(* IEC 61131-3 sources: SafePLC-Gen-Evaluation/Evaluation Results/butane/run_04, 2 files *)

(* ---- io_declarations.st ---- *)
(* ==================================================  *)
(* PLC I/O Variable Declarations — CODESYS 3.5  *)
(* Generated by SafePLC-Gen Multimodal  *)
(* ==================================================  *)

VAR_GLOBAL
    (* --- Analog Inputs ---  *)
    TI_2909_Raw                  AT %IW0       : INT := 0;    (* TI-2909 — Temperature indicator on process inlet l  *)
    TI_2917_Raw                  AT %IW2       : INT := 0;    (* TI-2917 — Temperature indicator high-high (HH), fa  *)
    TT_2909_Raw                  AT %IW4       : INT := 0;    (* TT-2909 — Temperature transmitter on process line,  *)
    TT_2911_Raw                  AT %IW6       : INT := 0;    (* TT-2911 — Temperature transmitter on process outle  *)
    TT_2917_Raw                  AT %IW8       : INT := 0;    (* TT-2917 — Temperature transmitter on heating mediu  *)
    XI_2901A_Raw                 AT %IW10      : INT := 0;    (* XI-2901A — Status indicator AVAILABLE for motor/fan  *)
    XI_2901B_Raw                 AT %IW12      : INT := 0;    (* XI-2901B — Status indicator AVAILABLE for motor/fan  *)
    (* --- Analog Outputs ---  *)
    KV_2904_Out                  AT %QW0       : INT := 0;    (* KV-2904 — Actuated valve on inlet process line, fa  *)
    (* --- Digital Inputs ---  *)
    ESD_3200                     AT %IX0.0     : BOOL := FALSE;    (* ESD-3200 — Emergency shutdown device/input, appears  *)
    HS_2901A                     AT %IX0.1     : BOOL := FALSE;    (* HS-2901A — Hand switch for motor/fan A control. Pan  *)
    HS_2901A1                    AT %IX0.2     : BOOL := FALSE;    (* HS-2901A1 — Hand switch LOCAL/REMOTE selector for mo  *)
    HS_2901A2                    AT %IX0.3     : BOOL := FALSE;    (* HS-2901A2 — Hand switch STOP/START for motor A at MC  *)
    HS_2901B                     AT %IX0.4     : BOOL := FALSE;    (* HS-2901B — Hand switch for motor/fan B control. Pan  *)
    HS_2901B1                    AT %IX0.5     : BOOL := FALSE;    (* HS-2901B1 — Hand switch LOCAL/REMOTE selector for mo  *)
    HS_2901B2                    AT %IX0.6     : BOOL := FALSE;    (* HS-2901B2 — Hand switch STOP/START for motor B at MC  *)
    HS_EMERGENCY_STOP_A_2901A    AT %IX0.7     : BOOL := FALSE;    (* HS-EMERGENCY-STOP-A-2901A — Emergency stop hand switch for motor A,   *)
    HS_EMERGENCY_STOP_B_2901B    AT %IX1.0     : BOOL := FALSE;    (* HS-EMERGENCY-STOP-B-2901B — Emergency stop hand switch for motor B,   *)
    HS_START_STOP_A_2901A        AT %IX1.1     : BOOL := FALSE;    (* HS-START-STOP-A-2901A — Field/local hand switch START/STOP for m  *)
    HS_START_STOP_B_2901B        AT %IX1.2     : BOOL := FALSE;    (* HS-START-STOP-B-2901B — Field/local hand switch START/STOP for m  *)
    PSD_2917                     AT %IX1.3     : BOOL := FALSE;    (* PSD-2917 — Pressure/Temperature shutdown device (PS  *)
    VSHH_2901A                   AT %IX1.4     : BOOL := FALSE;    (* VSHH-2901A — Vibration switch high-high on fan/motor   *)
    VSHH_2901B                   AT %IX1.5     : BOOL := FALSE;    (* VSHH-2901B — Vibration switch high-high on fan/motor   *)
END_VAR

(* ---- generated_code.st ---- *)
(* Generated by SafePLC-Gen Multimodal — CODESYS 3.5 *)
(* IEC 61131-3 Structured Text *)
(* Date: 2026-04-25T12:15:34.199960 *)

PROGRAM PRG_Compressor_2901

VAR
    TI_2909_Raw                  AT %IW0       : INT := 0;
    TI_2917_Raw                  AT %IW2       : INT := 0;
    TT_2909_Raw                  AT %IW4       : INT := 0;
    TT_2911_Raw                  AT %IW6       : INT := 0;
    TT_2917_Raw                  AT %IW8       : INT := 0;
    XI_2901A_Raw                 AT %IW10      : INT := 0;
    XI_2901B_Raw                 AT %IW12      : INT := 0;
    KV_2904_Out                  AT %QW0       : INT := 0;
    ESD_3200                     AT %IX0.0     : BOOL := FALSE;
    HS_2901A                     AT %IX0.1     : BOOL := FALSE;
    HS_2901A1                    AT %IX0.2     : BOOL := FALSE;
    HS_2901A2                    AT %IX0.3     : BOOL := FALSE;
    HS_2901B                     AT %IX0.4     : BOOL := FALSE;
    HS_2901B1                    AT %IX0.5     : BOOL := FALSE;
    HS_2901B2                    AT %IX0.6     : BOOL := FALSE;
    HS_EMERGENCY_STOP_A_2901A    AT %IX0.7     : BOOL := FALSE;
    HS_EMERGENCY_STOP_B_2901B    AT %IX1.0     : BOOL := FALSE;
    HS_START_STOP_A_2901A        AT %IX1.1     : BOOL := FALSE;
    HS_START_STOP_B_2901B        AT %IX1.2     : BOOL := FALSE;
    PSD_2917                     AT %IX1.3     : BOOL := FALSE;
    VSHH_2901A                   AT %IX1.4     : BOOL := FALSE;
    VSHH_2901B                   AT %IX1.5     : BOOL := FALSE;
    ESTOP                        AT %IX2.0     : BOOL := FALSE;
    MANUAL_RESET                 AT %IX2.1     : BOOL := FALSE;
    MCC_A_Out                    AT %QX0.0     : BOOL := FALSE;
    MCC_B_Out                    AT %QX0.1     : BOOL := FALSE;
    PSD_2917_Out                 AT %QX0.2     : BOOL := FALSE;
    MCC_A_and_MCC_B_Out          AT %QX0.3     : BOOL := FALSE;
END_VAR

VAR
    TI_2909_Scaled               : REAL := 0.0;
    TT_2909_Scaled               : REAL := 0.0;
    TT_2911_Scaled               : REAL := 0.0;
    TT_2917_Scaled               : REAL := 0.0;
    TI_2917_Scaled               : REAL := 0.0;
    XI_2901A_Scaled              : REAL := 0.0;
    XI_2901B_Scaled              : REAL := 0.0;

    TI_2909_HH_SP                : REAL := 120.0;
    TI_2909_H_SP                 : REAL := 110.0;
    TI_2909_L_SP                 : REAL := 10.0;
    TI_2909_LL_SP                : REAL := 5.0;
    TI_2909_Deadband             : REAL := 2.0;
    TI_2909_HH                   : BOOL := FALSE;
    TI_2909_H                    : BOOL := FALSE;
    TI_2909_L                    : BOOL := FALSE;
    TI_2909_LL                   : BOOL := FALSE;
    TI_2909_HH_Latch             : SR := (S1 := FALSE, R := FALSE, Q1 := FALSE);
    TI_2909_LL_Latch             : SR := (S1 := FALSE, R := FALSE, Q1 := FALSE);
    TI_2909_HH_Ack               : BOOL := FALSE;
    TI_2909_LL_Ack               : BOOL := FALSE;

    TT_2909_HH_SP                : REAL := 120.0;
    TT_2909_H_SP                 : REAL := 110.0;
    TT_2909_L_SP                 : REAL := 10.0;
    TT_2909_LL_SP                : REAL := 5.0;
    TT_2909_Deadband             : REAL := 2.0;
    TT_2909_HH                   : BOOL := FALSE;
    TT_2909_H                    : BOOL := FALSE;
    TT_2909_L                    : BOOL := FALSE;
    TT_2909_LL                   : BOOL := FALSE;
    TT_2909_HH_Latch             : SR := (S1 := FALSE, R := FALSE, Q1 := FALSE);
    TT_2909_LL_Latch             : SR := (S1 := FALSE, R := FALSE, Q1 := FALSE);
    TT_2909_HH_Ack               : BOOL := FALSE;
    TT_2909_LL_Ack               : BOOL := FALSE;

    TT_2911_HH_SP                : REAL := 120.0;
    TT_2911_H_SP                 : REAL := 110.0;
    TT_2911_L_SP                 : REAL := 10.0;
    TT_2911_LL_SP                : REAL := 5.0;
    TT_2911_Deadband             : REAL := 2.0;
    TT_2911_HH                   : BOOL := FALSE;
    TT_2911_H                    : BOOL := FALSE;
    TT_2911_L                    : BOOL := FALSE;
    TT_2911_LL                   : BOOL := FALSE;
    TT_2911_HH_Latch             : SR := (S1 := FALSE, R := FALSE, Q1 := FALSE);
    TT_2911_LL_Latch             : SR := (S1 := FALSE, R := FALSE, Q1 := FALSE);
    TT_2911_HH_Ack               : BOOL := FALSE;
    TT_2911_LL_Ack               : BOOL := FALSE;

    TIC_2911_SP                  : REAL := 60.0;
    TIC_2911_Kp                  : REAL := 1.5;
    TIC_2911_Ki                  : REAL := 0.05;
    TIC_2911_Error               : REAL := 0.0;
    TIC_2911_Integral            : REAL := 0.0;
    TIC_2911_Output              : REAL := 0.0;

    TT_2917_HH_SP                : REAL := 130.0;
    TT_2917_H_SP                 : REAL := 120.0;
    TT_2917_L_SP                 : REAL := 10.0;
    TT_2917_LL_SP                : REAL := 5.0;
    TT_2917_Deadband             : REAL := 2.0;
    TT_2917_HH                   : BOOL := FALSE;
    TT_2917_H                    : BOOL := FALSE;
    TT_2917_L                    : BOOL := FALSE;
    TT_2917_LL                   : BOOL := FALSE;
    TT_2917_HH_Latch             : SR := (S1 := FALSE, R := FALSE, Q1 := FALSE);
    TT_2917_LL_Latch             : SR := (S1 := FALSE, R := FALSE, Q1 := FALSE);
    TT_2917_HH_Ack               : BOOL := FALSE;
    TT_2917_LL_Ack               : BOOL := FALSE;

    TI_2917_HH_SP                : REAL := 130.0;
    TI_2917_H_SP                 : REAL := 120.0;
    TI_2917_L_SP                 : REAL := 10.0;
    TI_2917_LL_SP                : REAL := 5.0;
    TI_2917_Deadband             : REAL := 2.0;
    TI_2917_HH                   : BOOL := FALSE;
    TI_2917_H                    : BOOL := FALSE;
    TI_2917_L                    : BOOL := FALSE;
    TI_2917_LL                   : BOOL := FALSE;
    TI_2917_HH_Latch             : SR := (S1 := FALSE, R := FALSE, Q1 := FALSE);
    TI_2917_LL_Latch             : SR := (S1 := FALSE, R := FALSE, Q1 := FALSE);
    TI_2917_HH_Ack               : BOOL := FALSE;
    TI_2917_LL_Ack               : BOOL := FALSE;

    XI_2901A_HH_SP               : REAL := 90.0;
    XI_2901A_H_SP                : REAL := 80.0;
    XI_2901A_L_SP                : REAL := 10.0;
    XI_2901A_LL_SP               : REAL := 5.0;
    XI_2901A_Deadband            : REAL := 2.0;
    XI_2901A_HH                  : BOOL := FALSE;
    XI_2901A_H                   : BOOL := FALSE;
    XI_2901A_L                   : BOOL := FALSE;
    XI_2901A_LL                  : BOOL := FALSE;
    XI_2901A_HH_Latch            : SR := (S1 := FALSE, R := FALSE, Q1 := FALSE);
    XI_2901A_LL_Latch            : SR := (S1 := FALSE, R := FALSE, Q1 := FALSE);
    XI_2901A_HH_Ack              : BOOL := FALSE;
    XI_2901A_LL_Ack              : BOOL := FALSE;

    XI_2901B_HH_SP               : REAL := 90.0;
    XI_2901B_H_SP                : REAL := 80.0;
    XI_2901B_L_SP                : REAL := 10.0;
    XI_2901B_LL_SP               : REAL := 5.0;
    XI_2901B_Deadband            : REAL := 2.0;
    XI_2901B_HH                  : BOOL := FALSE;
    XI_2901B_H                   : BOOL := FALSE;
    XI_2901B_L                   : BOOL := FALSE;
    XI_2901B_LL                  : BOOL := FALSE;
    XI_2901B_HH_Latch            : SR := (S1 := FALSE, R := FALSE, Q1 := FALSE);
    XI_2901B_LL_Latch            : SR := (S1 := FALSE, R := FALSE, Q1 := FALSE);
    XI_2901B_HH_Ack              : BOOL := FALSE;
    XI_2901B_LL_Ack              : BOOL := FALSE;

    LOOP_2917_TRIP               : BOOL := FALSE;
    LOOP_2901A_TRIP              : BOOL := FALSE;
    LOOP_2901B_TRIP              : BOOL := FALSE;
    LOOP_3200_TRIP               : BOOL := FALSE;

    TT_2917_HH_Trip              : BOOL := FALSE;
    TT_2917_LL_Trip              : BOOL := FALSE;
    VSHH_2901A_HH                : BOOL := FALSE;
    VSHH_2901A_LL                : BOOL := FALSE;
    VSHH_2901B_HH                : BOOL := FALSE;
    VSHH_2901B_LL                : BOOL := FALSE;
    ESD_3200_HH                  : BOOL := FALSE;
    ESD_3200_LL                  : BOOL := FALSE;

    SAFE_STATE                   : BOOL := FALSE;

    MotorA_LocalMode             : BOOL := FALSE;
    MotorA_StartCmd              : BOOL := FALSE;
    MotorA_StopCmd               : BOOL := FALSE;
    MotorA_Run                   : BOOL := FALSE;
    MotorA_Latch                 : SR := (S1 := FALSE, R := FALSE, Q1 := FALSE);

    MotorB_LocalMode             : BOOL := FALSE;
    MotorB_StartCmd              : BOOL := FALSE;
    MotorB_StopCmd               : BOOL := FALSE;
    MotorB_Run                   : BOOL := FALSE;
    MotorB_Latch                 : SR := (S1 := FALSE, R := FALSE, Q1 := FALSE);

    StartupDelay                 : TON := (IN := FALSE, PT := T#3S);

    System_Alarm                 : BOOL := FALSE;
    FirstScan                    : BOOL := TRUE;
END_VAR

IF FirstScan THEN
    LOOP_2917_TRIP       := TRUE;
    LOOP_2901A_TRIP      := TRUE;
    LOOP_2901B_TRIP      := TRUE;
    LOOP_3200_TRIP       := TRUE;
    SAFE_STATE           := TRUE;
    KV_2904_Out          := 6554;
    MCC_A_Out            := FALSE;
    MCC_B_Out            := FALSE;
    PSD_2917_Out         := FALSE;
    MCC_A_and_MCC_B_Out  := FALSE;
    TIC_2911_Integral    := 0.0;
    FirstScan            := FALSE;
    RETURN;
END_IF;

TI_2909_Scaled  := ((INT_TO_REAL(TI_2909_Raw)  - 6554.0) / (32767.0 - 6554.0)) * 150.0;
TT_2909_Scaled  := ((INT_TO_REAL(TT_2909_Raw)  - 6554.0) / (32767.0 - 6554.0)) * 150.0;
TT_2911_Scaled  := ((INT_TO_REAL(TT_2911_Raw)  - 6554.0) / (32767.0 - 6554.0)) * 150.0;
TT_2917_Scaled  := ((INT_TO_REAL(TT_2917_Raw)  - 6554.0) / (32767.0 - 6554.0)) * 150.0;
TI_2917_Scaled  := ((INT_TO_REAL(TI_2917_Raw)  - 6554.0) / (32767.0 - 6554.0)) * 150.0;
XI_2901A_Scaled := ((INT_TO_REAL(XI_2901A_Raw) - 6554.0) / (32767.0 - 6554.0)) * 100.0;
XI_2901B_Scaled := ((INT_TO_REAL(XI_2901B_Raw) - 6554.0) / (32767.0 - 6554.0)) * 100.0;

TT_2917_HH_Trip := TT_2917_Scaled >= TT_2917_HH_SP;
TT_2917_LL_Trip := TT_2917_Scaled <= TT_2917_LL_SP;
VSHH_2901A_HH   := VSHH_2901A;
VSHH_2901A_LL   := FALSE;
VSHH_2901B_HH   := VSHH_2901B;
VSHH_2901B_LL   := FALSE;
ESD_3200_HH     := ESD_3200;
ESD_3200_LL     := FALSE;

IF TT_2917_HH_Trip OR TT_2917_LL_Trip OR PSD_2917 THEN
    LOOP_2917_TRIP := TRUE;
ELSIF LOOP_2917_TRIP AND MANUAL_RESET
      AND NOT TT_2917_HH_Trip AND NOT TT_2917_LL_Trip AND NOT PSD_2917 THEN
    LOOP_2917_TRIP := FALSE;
END_IF;

IF VSHH_2901A_HH OR VSHH_2901A_LL OR HS_EMERGENCY_STOP_A_2901A THEN
    LOOP_2901A_TRIP := TRUE;
ELSIF LOOP_2901A_TRIP AND MANUAL_RESET
      AND NOT VSHH_2901A_HH AND NOT VSHH_2901A_LL AND NOT HS_EMERGENCY_STOP_A_2901A THEN
    LOOP_2901A_TRIP := FALSE;
END_IF;

IF VSHH_2901B_HH OR VSHH_2901B_LL OR HS_EMERGENCY_STOP_B_2901B THEN
    LOOP_2901B_TRIP := TRUE;
ELSIF LOOP_2901B_TRIP AND MANUAL_RESET
      AND NOT VSHH_2901B_HH AND NOT VSHH_2901B_LL AND NOT HS_EMERGENCY_STOP_B_2901B THEN
    LOOP_2901B_TRIP := FALSE;
END_IF;

IF ESD_3200_HH OR ESD_3200_LL THEN
    LOOP_3200_TRIP := TRUE;
ELSIF LOOP_3200_TRIP AND MANUAL_RESET
      AND NOT ESD_3200_HH AND NOT ESD_3200_LL THEN
    LOOP_3200_TRIP := FALSE;
END_IF;

SAFE_STATE := ESTOP
              OR LOOP_2917_TRIP
              OR LOOP_2901A_TRIP
              OR LOOP_2901B_TRIP
              OR LOOP_3200_TRIP;

IF NOT SAFE_STATE THEN
    TIC_2911_Error    := TIC_2911_SP - TT_2911_Scaled;
    TIC_2911_Integral := TIC_2911_Integral + (TIC_2911_Ki * TIC_2911_Error);
    IF TIC_2911_Integral > 100.0 THEN
        TIC_2911_Integral := 100.0;
    ELSIF TIC_2911_Integral < 0.0 THEN
        TIC_2911_Integral := 0.0;
    END_IF;
    TIC_2911_Output := (TIC_2911_Kp * TIC_2911_Error) + TIC_2911_Integral;
    IF TIC_2911_Output > 100.0 THEN
        TIC_2911_Output := 100.0;
    ELSIF TIC_2911_Output < 0.0 THEN
        TIC_2911_Output := 0.0;
    END_IF;
    KV_2904_Out := REAL_TO_INT(6554.0 + (TIC_2911_Output / 100.0) * (32767.0 - 6554.0));

    MotorA_LocalMode := HS_2901A1;
    IF MotorA_LocalMode THEN
        MotorA_StartCmd := HS_START_STOP_A_2901A;
        MotorA_StopCmd  := NOT HS_START_STOP_A_2901A;
    ELSE
        MotorA_StartCmd := HS_2901A AND HS_2901A2;
        MotorA_StopCmd  := NOT HS_2901A2;
    END_IF;
    MotorA_Latch(S1 := MotorA_StartCmd, R := MotorA_StopCmd);
    MotorA_Run := MotorA_Latch.Q1;

    MotorB_LocalMode := HS_2901B1;
    IF MotorB_LocalMode THEN
        MotorB_StartCmd := HS_START_STOP_B_2901B;
        MotorB_StopCmd  := NOT HS_START_STOP_B_2901B;
    ELSE
        MotorB_StartCmd := HS_2901B AND HS_2901B2;
        MotorB_StopCmd  := NOT HS_2901B2;
    END_IF;
    MotorB_Latch(S1 := MotorB_StartCmd, R := MotorB_StopCmd);
    MotorB_Run := MotorB_Latch.Q1;

    StartupDelay(IN := MotorA_Run OR MotorB_Run, PT := T#3S);

    MCC_A_Out           := MotorA_Run AND StartupDelay.Q;
    MCC_B_Out           := MotorB_Run AND StartupDelay.Q;
    PSD_2917_Out        := TRUE;
    MCC_A_and_MCC_B_Out := MCC_A_Out AND MCC_B_Out;
ELSE
    KV_2904_Out         := 6554;
    MCC_A_Out           := FALSE;
    MCC_B_Out           := FALSE;
    PSD_2917_Out        := FALSE;
    MCC_A_and_MCC_B_Out := FALSE;
    TIC_2911_Integral   := 0.0;
END_IF;

(* TI_2909 four-level alarms *)
IF TI_2909_Scaled >= TI_2909_HH_SP THEN
    TI_2909_HH_Latch.S1 := TRUE;
ELSIF TI_2909_Scaled <= (TI_2909_HH_SP - TI_2909_Deadband) THEN
    TI_2909_HH_Latch.S1 := FALSE;
END_IF;
TI_2909_HH_Latch(S1 := TI_2909_HH_Latch.S1, R := TI_2909_HH_Ack AND (TI_2909_Scaled < TI_2909_HH_SP));
TI_2909_HH := TI_2909_HH_Latch.Q1;
TI_2909_H  := TI_2909_Scaled >= TI_2909_H_SP AND TI_2909_Scaled < TI_2909_HH_SP;
TI_2909_L  := TI_2909_Scaled <= TI_2909_L_SP AND TI_2909_Scaled > TI_2909_LL_SP;
IF TI_2909_Scaled <= TI_2909_LL_SP THEN
    TI_2909_LL_Latch.S1 := TRUE;
ELSIF TI_2909_Scaled >= (TI_2909_LL_SP + TI_2909_Deadband) THEN
    TI_2909_LL_Latch.S1 := FALSE;
END_IF;
TI_2909_LL_Latch(S1 := TI_2909_LL_Latch.S1, R := TI_2909_LL_Ack AND (TI_2909_Scaled > TI_2909_LL_SP));
TI_2909_LL := TI_2909_LL_Latch.Q1;

(* TT_2909 four-level alarms *)
IF TT_2909_Scaled >= TT_2909_HH_SP THEN
    TT_2909_HH_Latch.S1 := TRUE;
ELSIF TT_2909_Scaled <= (TT_2909_HH_SP - TT_2909_Deadband) THEN
    TT_2909_HH_Latch.S1 := FALSE;
END_IF;
TT_2909_HH_Latch(S1 := TT_2909_HH_Latch.S1, R := TT_2909_HH_Ack AND (TT_2909_Scaled < TT_2909_HH_SP));
TT_2909_HH := TT_2909_HH_Latch.Q1;
TT_2909_H  := TT_2909_Scaled >= TT_2909_H_SP AND TT_2909_Scaled < TT_2909_HH_SP;
TT_2909_L  := TT_2909_Scaled <= TT_2909_L_SP AND TT_2909_Scaled > TT_2909_LL_SP;
IF TT_2909_Scaled <= TT_2909_LL_SP THEN
    TT_2909_LL_Latch.S1 := TRUE;
ELSIF TT_2909_Scaled >= (TT_2909_LL_SP + TT_2909_Deadband) THEN
    TT_2909_LL_Latch.S1 := FALSE;
END_IF;
TT_2909_LL_Latch(S1 := TT_2909_LL_Latch.S1, R := TT_2909_LL_Ack AND (TT_2909_Scaled > TT_2909_LL_SP));
TT_2909_LL := TT_2909_LL_Latch.Q1;

(* TT_2911 four-level alarms *)
IF TT_2911_Scaled >= TT_2911_HH_SP THEN
    TT_2911_HH_Latch.S1 := TRUE;
ELSIF TT_2911_Scaled <= (TT_2911_HH_SP - TT_2911_Deadband) THEN
    TT_2911_HH_Latch.S1 := FALSE;
END_IF;
TT_2911_HH_Latch(S1 := TT_2911_HH_Latch.S1, R := TT_2911_HH_Ack AND (TT_2911_Scaled < TT_2911_HH_SP));
TT_2911_HH := TT_2911_HH_Latch.Q1;
TT_2911_H  := TT_2911_Scaled >= TT_2911_H_SP AND TT_2911_Scaled < TT_2911_HH_SP;
TT_2911_L  := TT_2911_Scaled <= TT_2911_L_SP AND TT_2911_Scaled > TT_2911_LL_SP;
IF TT_2911_Scaled <= TT_2911_LL_SP THEN
    TT_2911_LL_Latch.S1 := TRUE;
ELSIF TT_2911_Scaled >= (TT_2911_LL_SP + TT_2911_Deadband) THEN
    TT_2911_LL_Latch.S1 := FALSE;
END_IF;
TT_2911_LL_Latch(S1 := TT_2911_LL_Latch.S1, R := TT_2911_LL_Ack AND (TT_2911_Scaled > TT_2911_LL_SP));
TT_2911_LL := TT_2911_LL_Latch.Q1;

(* TT_2917 four-level alarms *)
IF TT_2917_Scaled >= TT_2917_HH_SP THEN
    TT_2917_HH_Latch.S1 := TRUE;
ELSIF TT_2917_Scaled <= (TT_2917_HH_SP - TT_2917_Deadband) THEN
    TT_2917_HH_Latch.S1 := FALSE;
END_IF;
TT_2917_HH_Latch(S1 := TT_2917_HH_Latch.S1, R := TT_2917_HH_Ack AND (TT_2917_Scaled < TT_2917_HH_SP));
TT_2917_HH := TT_2917_HH_Latch.Q1;
TT_2917_H  := TT_2917_Scaled >= TT_2917_H_SP AND TT_2917_Scaled < TT_2917_HH_SP;
TT_2917_L  := TT_2917_Scaled <= TT_2917_L_SP AND TT_2917_Scaled > TT_2917_LL_SP;
IF TT_2917_Scaled <= TT_2917_LL_SP THEN
    TT_2917_LL_Latch.S1 := TRUE;
ELSIF TT_2917_Scaled >= (TT_2917_LL_SP + TT_2917_Deadband) THEN
    TT_2917_LL_Latch.S1 := FALSE;
END_IF;
TT_2917_LL_Latch(S1 := TT_2917_LL_Latch.S1, R := TT_2917_LL_Ack AND (TT_2917_Scaled > TT_2917_LL_SP));
TT_2917_LL := TT_2917_LL_Latch.Q1;

(* TI_2917 four-level alarms *)
IF TI_2917_Scaled >= TI_2917_HH_SP THEN
    TI_2917_HH_Latch.S1 := TRUE;
ELSIF TI_2917_Scaled <= (TI_2917_HH_SP - TI_2917_Deadband) THEN
    TI_2917_HH_Latch.S1 := FALSE;
END_IF;
TI_2917_HH_Latch(S1 := TI_2917_HH_Latch.S1, R := TI_2917_HH_Ack AND (TI_2917_Scaled < TI_2917_HH_SP));
TI_2917_HH := TI_2917_HH_Latch.Q1;
TI_2917_H  := TI_2917_Scaled >= TI_2917_H_SP AND TI_2917_Scaled < TI_2917_HH_SP;
TI_2917_L  := TI_2917_Scaled <= TI_2917_L_SP AND TI_2917_Scaled > TI_2917_LL_SP;
IF TI_2917_Scaled <= TI_2917_LL_SP THEN
    TI_2917_LL_Latch.S1 := TRUE;
ELSIF TI_2917_Scaled >= (TI_2917_LL_SP + TI_2917_Deadband) THEN
    TI_2917_LL_Latch.S1 := FALSE;
END_IF;
TI_2917_LL_Latch(S1 := TI_2917_LL_Latch.S1, R := TI_2917_LL_Ack AND (TI_2917_Scaled > TI_2917_LL_SP));
TI_2917_LL := TI_2917_LL_Latch.Q1;

(* XI_2901A four-level alarms *)
IF XI_2901A_Scaled >= XI_2901A_HH_SP THEN
    XI_2901A_HH_Latch.S1 := TRUE;
ELSIF XI_2901A_Scaled <= (XI_2901A_HH_SP - XI_2901A_Deadband) THEN
    XI_2901A_HH_Latch.S1 := FALSE;
END_IF;
XI_2901A_HH_Latch(S1 := XI_2901A_HH_Latch.S1, R := XI_2901A_HH_Ack AND (XI_2901A_Scaled < XI_2901A_HH_SP));
XI_2901A_HH := XI_2901A_HH_Latch.Q1;
XI_2901A_H  := XI_2901A_Scaled >= XI_2901A_H_SP AND XI_2901A_Scaled < XI_2901A_HH_SP;
XI_2901A_L  := XI_2901A_Scaled <= XI_2901A_L_SP AND XI_2901A_Scaled > XI_2901A_LL_SP;
IF XI_2901A_Scaled <= XI_2901A_LL_SP THEN
    XI_2901A_LL_Latch.S1 := TRUE;
ELSIF XI_2901A_Scaled >= (XI_2901A_LL_SP + XI_2901A_Deadband) THEN
    XI_2901A_LL_Latch.S1 := FALSE;
END_IF;
XI_2901A_LL_Latch(S1 := XI_2901A_LL_Latch.S1, R := XI_2901A_LL_Ack AND (XI_2901A_Scaled > XI_2901A_LL_SP));
XI_2901A_LL := XI_2901A_LL_Latch.Q1;

(* XI_2901B four-level alarms *)
IF XI_2901B_Scaled >= XI_2901B_HH_SP THEN
    XI_2901B_HH_Latch.S1 := TRUE;
ELSIF XI_2901B_Scaled <= (XI_2901B_HH_SP - XI_2901B_Deadband) THEN
    XI_2901B_HH_Latch.S1 := FALSE;
END_IF;
XI_2901B_HH_Latch(S1 := XI_2901B_HH_Latch.S1, R := XI_2901B_HH_Ack AND (XI_2901B_Scaled < XI_2901B_HH_SP));
XI_2901B_HH := XI_2901B_HH_Latch.Q1;
XI_2901B_H  := XI_2901B_Scaled >= XI_2901B_H_SP AND XI_2901B_Scaled < XI_2901B_HH_SP;
XI_2901B_L  := XI_2901B_Scaled <= XI_2901B_L_SP AND XI_2901B_Scaled > XI_2901B_LL_SP;
IF XI_2901B_Scaled <= XI_2901B_LL_SP THEN
    XI_2901B_LL_Latch.S1 := TRUE;
ELSIF XI_2901B_Scaled >= (XI_2901B_LL_SP + XI_2901B_Deadband) THEN
    XI_2901B_LL_Latch.S1 := FALSE;
END_IF;
XI_2901B_LL_Latch(S1 := XI_2901B_LL_Latch.S1, R := XI_2901B_LL_Ack AND (XI_2901B_Scaled > XI_2901B_LL_SP));
XI_2901B_LL := XI_2901B_LL_Latch.Q1;

System_Alarm :=
    TI_2909_HH_Latch.Q1 OR TI_2909_LL_Latch.Q1 OR TI_2909_H OR TI_2909_L OR
    TT_2909_HH_Latch.Q1 OR TT_2909_LL_Latch.Q1 OR TT_2909_H OR TT_2909_L OR
    TT_2911_HH_Latch.Q1 OR TT_2911_LL_Latch.Q1 OR TT_2911_H OR TT_2911_L OR
    TT_2917_HH_Latch.Q1 OR TT_2917_LL_Latch.Q1 OR TT_2917_H OR TT_2917_L OR
    TI_2917_HH_Latch.Q1 OR TI_2917_LL_Latch.Q1 OR TI_2917_H OR TI_2917_L OR
    XI_2901A_HH_Latch.Q1 OR XI_2901A_LL_Latch.Q1 OR XI_2901A_H OR XI_2901A_L OR
    XI_2901B_HH_Latch.Q1 OR XI_2901B_LL_Latch.Q1 OR XI_2901B_H OR XI_2901B_L OR
    SAFE_STATE;

END_PROGRAM
